TYPE ST_NCTOPLC :
STRUCT
	(* SDS *)
	stBaseDevice				:ST_BaseDeviceIn;

	(* SD6/SC6/SI6 *)
	stCIA402						:ST_CIA402In;

END_STRUCT
END_TYPE

(* stored: Version 1.1.0.1, ProductVersion 3.1.4024.15
   DUT ST_NCTOPLC: Id {f9474bc7-6220-4c63-b8b6-7c0614611969} *)
